(* IEC 61131-3 sources: codesys-framework/txt/application/WeVe Core (library)/60 Event/FB_EventGroup, 8 files *)

(* ---- Condition.method.st ---- *)
// Doorgeefluik naar I_Event.Condition van event iEvent (enum van de eigenaar).
// Geeft Active van dat event terug, FALSE bij een ongeldige index.
METHOD Condition : BOOL
VAR_INPUT
	iEvent 			: INT;
	xCondition 		: BOOL;
	scPayload 		: SC_EventPayload := (asPayload := [10('')]);	// mag weggelaten worden
END_VAR
VAR
	fbEvent 		: I_Event;
END_VAR

// --- BEGIN IMPLEMENTATION ---

fbEvent := GetEvent(iEvent);

IF fbEvent = 0 THEN
	Condition := FALSE;
	RETURN;
END_IF

Condition := fbEvent.Condition(xCondition := xCondition, scPayload := scPayload);

(* ---- FB_Init.method.st ---- *)
//FB_Init is always available implicitly and it is used primarily for initialization.
//The return value is not evaluated. For a specific influence, you can also declare the
//methods explicitly and provide additional code there with the standard initialization
//code. You can evaluate the return value.
METHOD FB_Init: BOOL
VAR_INPUT
    bInitRetains: BOOL; // TRUE: the retain variables are initialized (reset warm / reset cold)
    bInCopyCode: BOOL;  // TRUE: the instance will be copied to the copy code afterward (online change)

	fbLogger 			: I_Logger;		// mag 0 zijn: events houden dan enkel hun toestand bij
	nSubMachine 		: USINT;		// bron van alle events van deze groep
	nSubMachineId 		: USINT;
END_VAR

// --- BEGIN IMPLEMENTATION ---

// Enkel referenties en waarden bewaren, geen methodes aanroepen
_fbLogger 		:= fbLogger;
_nSubMachine 	:= nSubMachine;
_nSubMachineId 	:= nSubMachineId;

(* ---- GetEvent.method.st ---- *)
// Door de afgeleide groep: event iEvent teruggeven, 0 bij een ongeldige index.
//   IF iEvent >= 0 AND iEvent < Count THEN
//       GetEvent := _afbEvents[iEvent];
//   ELSE
//       GetEvent := 0;
//   END_IF
METHOD ABSTRACT GetEvent : I_Event
VAR_INPUT
	iEvent 			: INT;
END_VAR

(* ---- HasAlarm.prop.st ---- *)
// Alarm = level Operator of Supervisor. EventIsAlarm_OnlyLogLevel telt niet mee: wordt enkel gelogd.
PROPERTY HasAlarm : BOOL
// --- BEGIN IMPLEMENTATION ---

// ----------- GET -----------
VAR
	i 			: INT;
	fbEvent 	: I_Event;
END_VAR

// -- BEGIN IMPLEMENTATION GET --
HasAlarm := FALSE;

FOR i := 0 TO Count - 1 DO
	fbEvent := GetEvent(i);
	IF fbEvent <> 0 THEN
		IF fbEvent.Active AND (fbEvent.Level = E_EventLevels.EventIsAlarm_OperatorLevel OR fbEvent.Level = E_EventLevels.EventIsAlarm_SupervisorLevel) THEN
			HasAlarm := TRUE;
			RETURN;
		END_IF
	END_IF
END_FOR

(* ---- HasWarning.prop.st ---- *)
PROPERTY HasWarning : BOOL
// --- BEGIN IMPLEMENTATION ---

// ----------- GET -----------
VAR
	i 			: INT;
	fbEvent 	: I_Event;
END_VAR

// -- BEGIN IMPLEMENTATION GET --
HasWarning := FALSE;

FOR i := 0 TO Count - 1 DO
	fbEvent := GetEvent(i);
	IF fbEvent <> 0 THEN
		IF fbEvent.Active AND (fbEvent.Level = E_EventLevels.EventIsWarning_NotUrgent OR fbEvent.Level = E_EventLevels.EventIsWarning_Urgent) THEN
			HasWarning := TRUE;
			RETURN;
		END_IF
	END_IF
END_FOR

(* ---- Initialize.method.st ---- *)
// Eenmalig bij de opstart: logger doorgeven aan alle events en hun config invullen.
// Mag meermaals aangeroepen worden, enkel de eerste keer doet iets.
// TRUE = klaar.
METHOD Initialize : BOOL
VAR_INPUT
END_VAR
VAR
	i 			: INT;
	fbEvent 	: I_Event;
END_VAR

// --- BEGIN IMPLEMENTATION ---

IF _xInitialized THEN
	Initialize := TRUE;
	RETURN;
END_IF

FOR i := 0 TO Count - 1 DO
	fbEvent := GetEvent(i);
	IF fbEvent <> 0 THEN
		fbEvent.Logger := _fbLogger;
	END_IF
END_FOR

ConfigureEvents();

_xInitialized := TRUE;
Initialize := TRUE;

(* ---- Log.method.st ---- *)
// Doorgeefluik naar I_Event.Log van event iEvent (enum van de eigenaar).
// FALSE bij een ongeldige index.
METHOD Log : BOOL
VAR_INPUT
	iEvent 			: INT;
	scPayload 		: SC_EventPayload := (asPayload := [10('')]);	// mag weggelaten worden
END_VAR
VAR
	fbEvent 		: I_Event;
END_VAR

// --- BEGIN IMPLEMENTATION ---

fbEvent := GetEvent(iEvent);

IF fbEvent = 0 THEN
	Log := FALSE;
	RETURN;
END_IF

Log := fbEvent.Log(scPayload := scPayload);

(* ---- Reset.method.st ---- *)
// Reset alle events van de groep. Elk event beslist zelf of het mag (conditie weg).
// TRUE = geen enkel event nog actief.
METHOD Reset : BOOL
VAR_INPUT
END_VAR
VAR
	i 			: INT;
	fbEvent 	: I_Event;
	xAllReset 	: BOOL := TRUE;
END_VAR

// --- BEGIN IMPLEMENTATION ---

FOR i := 0 TO Count - 1 DO
	fbEvent := GetEvent(i);
	IF fbEvent <> 0 THEN
		// Reset altijd aanroepen, ook als een vorig event al FALSE gaf
		IF NOT fbEvent.Reset() THEN
			xAllReset := FALSE;
		END_IF
	END_IF
END_FOR

Reset := xAllReset;
